FUNCTION_BLOCK FB_TwinSAFE
VAR_INPUT
	ES1_Restart: BOOL;
	ES2_Restart: BOOL;
	ES3_Restart: BOOL;
	ES4_Restart: BOOL;
END_VAR
VAR_OUTPUT
	outStateSafe: BOOL;
END_VAR
VAR
	rt_TSafe_OK: R_TRIG;
	rt_TSafe_Err: R_TRIG;
	ton_TSafe_OK: TON;
	ton_TSafe_Err_Reset_ON: TON;
	ton_TSafe_Err_Reset_OFF: TON;	
END_VAR
VAR_IN_OUT
	stTS: ST_TwinSAFE;
END_VAR

stTS.stSafetyOut.ES1_PB_Restart:=ES1_Restart;
stTS.stSafetyOut.ES2_PB_Restart:=ES2_Restart;
stTS.stSafetyOut.ES3_PB_Restart:=ES3_Restart;
stTS.stSafetyOut.ES4_PB_Restart:=ES4_Restart;


//stTS.TSafeOut.Restart:=ES1_Restart;

ton_TSafe_OK(IN:=stTS.TSafeIn.InRun AND NOT stTS.TSafeIn.COM_Err, PT:=T#1S );
IF ton_TSafe_OK.Q 
AND stTS.stSafetyIn.ES1_State
AND stTS.stSafetyIn.ES2_State
AND stTS.stSafetyIn.ES3_State
AND stTS.stSafetyIn.ES4_State
THEN;
	outStateSafe:=TRUE;
ELSE;
	outStateSafe:=FALSE;	
END_IF
rt_TSafe_OK(CLK:=ton_TSafe_OK.Q );
IF rt_TSafe_OK.Q THEN;
	//m_Print_Success_Message();
END_IF



rt_TSafe_Err(CLK:=stTS.TSafeIn.COM_Err);
IF rt_TSafe_Err.Q THEN;
	//m_Print_Error_Message();
END_IF

ton_TSafe_Err_Reset_ON(IN:=stTS.TSafeIn.COM_Err AND NOT stTS.TSafeOut.ErrACK, PT:=T#2S );
IF ton_TSafe_Err_Reset_ON.Q THEN;
	stTS.TSafeOut.ErrACK:=TRUE;
END_IF

ton_TSafe_Err_Reset_OFF(IN:=stTS.TSafeOut.ErrACK, PT:=T#1S );
IF ton_TSafe_Err_Reset_OFF.Q THEN;
	stTS.TSafeOut.ErrACK:=FALSE;
END_IF

METHOD m_Print_Error_Message : BOOL
VAR_INPUT
END_VAR

VAR
	i: INT;
	sActErrorID: STRING(11);
	sModuleDescription: STRING(80);
END_VAR

sActErrorID:='0x999x0';
sModuleDescription:='TwinSAFE Group';

FOR i:=100 TO 2 BY -1 DO
	Buffer_Act_Message[i]:=Buffer_Act_Message[i-1];
END_FOR

Buffer_Act_Message[1].sDateTime:=sRealTime_Date;
Buffer_Act_Message[1].sErrID:=sActErrorID;
Buffer_Act_Message[1].sModuleDescription:=sModuleDescription;
Buffer_Act_Message[1].sLevel:='Error';
Buffer_Act_Message[1].sErrorMessage:='';

Buffer_Act_Message[1].sErrorMessage:=CONCAT(Buffer_Act_Message[1].sErrorMessage,'TwinSAFE group has a communication error');
FUN_Write_Line_To_History();
END_METHOD

METHOD m_Print_Success_Message : BOOL
VAR_INPUT
END_VAR

VAR
	i: INT;
	sActErrorID: STRING(11);
	sModuleDescription: STRING(80);
END_VAR

sActErrorID:='0x999x0';
sModuleDescription:='TwinSAFE Group';

FOR i:=1000 TO 2 BY -1 DO
	Buffer_Act_History[i]:=Buffer_Act_History[i-1];
END_FOR

Buffer_Act_History[1].sDateTime:=sRealTime_Date;
Buffer_Act_History[1].sErrID:=sActErrorID;
Buffer_Act_History[1].sModuleDescription:=sModuleDescription;
Buffer_Act_History[1].sLevel:='Message';
Buffer_Act_History[1].sErrorMessage:='';

Buffer_Act_History[1].sErrorMessage:=CONCAT(Buffer_Act_History[1].sErrorMessage,'TwinSAFE state is OK');
END_METHOD

END_FUNCTION_BLOCK

(* stored: Version 1.1.0.1, ProductVersion 3.1.4024.13
   POU FB_TwinSAFE: Id {4ab5defe-eed2-490f-bb56-b846d8da8e90}, SpecialFunc None
   Method m_Print_Error_Message: Id {083c4f03-3c6b-4b7e-b608-334a475b1764}
   Method m_Print_Success_Message: Id {0548d864-a910-432c-b329-bfbcc1612a5d} *)
